(* IEC 61131-3 sources: 2026_Projet_YGO_ExcavatriceDragage/CODE_BACKUP/CODE_20260822_IntroductionTestCI/J_SUPERVISION/_TYPES/4_JOYSTICK_ACQUISITION, 9 files *)

(* ---- ST_AcquisitionInterPrg.st ---- *)
(* ═══════════════════════════════════════════════════════════════
   🧲 ST_AcquisitionInterPrg — Bus d'échange inter-PRG produit par PRG_02_Acquisition
   ───────────────────────────────────────────────────────────────
   🎯 Rôle : Encapsuler les mesures câbles/vitesses, les états joystick qualifiés,
      les positions M3 et les diagnostics DI publiés par PRG_02_Acquisition vers
      les consommateurs (PRG_03/04/05/07, FB_TroubleshootingView).
   📤 Producteur unique : PRG_02_Acquisition (VAR_OUTPUT Data : ST_AcquisitionInterPrg).
   📄 Doc : DOC/AF/AF_Partie-06_Acquisition_Qualification_IO_v2.3.md
   🔌 Architecture : Bus de données typé — encapsulation des échanges inter-PRG.
   ═══════════════════════════════════════════════════════════════ *)

TYPE ST_AcquisitionInterPrg :
STRUCT
    // === 🧲 Mesures câbles & vitesses treuils M1/M2 ===
    CablePosM1              : REAL; // 📏 Position cable M1 calibree (metres)
    CablePosM2              : REAL; // 📏 Position cable M2 calibree (metres)
    M1_Speed_Mps            : REAL; // 📏 Vitesse absolue M1 (m/s)
    M1_SignedSpeed_Mps      : REAL; // 📏 Vitesse signee M1 (+:Montee, -:Descente) (m/s)
    M1_SpeedValid           : BOOL; // 🟢 Validite mesure vitesse M1
    M2_Speed_Mps            : REAL; // 📏 Vitesse absolue M2 (m/s)
    M2_SignedSpeed_Mps      : REAL; // 📏 Vitesse signee M2 (+:Montee, -:Descente) (m/s)
    M2_SpeedValid           : BOOL; // 🟢 Validite mesure vitesse M2

    // === 🕹️ États joystick qualifiés ===
    JoystickDeadmanArmed    : BOOL; // 🔒 Homme-mort joystick arme (1=Arme)
    JoystickYNeutral        : BOOL; // 🟢 Axe Y joystick au neutre
    JoystickDirectionX      : INT;  // 🎯 Sens X demande (-1:Gauche, 0:Neutre, 1:Droite)
    JoystickSpeedPctX       : REAL; // 📈 Magnitude deviation axe X en % (0..100)
    JoystickXNeutral        : BOOL; // 🟢 Axe X joystick au neutre

    // === 🎯 Positions translation M3 (zones cumulatives + points exacts) ===
    TranslationPosTremie      : BOOL; // 📍 Zone Tremie (1=Present)
    TranslationPosPV          : BOOL; // 📍 Zone pre-ralentissement PV (1=Present)
    TranslationPosP2          : BOOL; // 📍 Zone P2 (1=Present)
    TranslationPosP1          : BOOL; // 📍 Zone P1 (1=Present)
    TranslationPosMaintenance : BOOL; // 📍 Zone Maintenance (1=Present)
    TranslationAtTremie       : BOOL; // 🎯 Position exacte Tremie (1=Atteint)
    TranslationAtPV           : BOOL; // 🎯 Position exacte PV (1=Atteint)
    TranslationAtP2           : BOOL; // 🎯 Position exacte P2 (1=Atteint)
    TranslationAtP1           : BOOL; // 🎯 Position exacte P1 (1=Atteint)
    TranslationAtMaintenance  : BOOL; // 🎯 Position exacte Maintenance (1=Atteint)
    M3_LimitSwitchFwd         : BOOL; // 🛡️ Fin de course avant M3 (1=Actionne)
    M3_LimitSwitchRev         : BOOL; // 🛡️ Fin de course arriere M3 (1=Actionne)
    M3_SensorWordIncoherent   : BOOL; // ❌ Incoherence detectee mot capteurs M3
    M3_SensorsWord             : BYTE; // 📊 Mot d'etat capteurs M3

    // === 🩺 Diagnostics modules DI & codeurs ===
    LocalDigitalIoOk         : BOOL; // 🟢 Module Local_Digital_IO OK
    Vh0800EndOk              : BOOL; // 🟢 Module VH_0800END OK
    Vh0808EtpOk              : BOOL; // 🟢 Module VH_0808ETP OK
    InputModuleFault         : BOOL; // ❌ Defaut sur au moins un module DI
    M1_EncoderIncoherent     : BOOL; // ❌ Mesure codeur M1 incoherente
    M2_EncoderIncoherent     : BOOL; // ❌ Mesure codeur M2 incoherente
    M1_EncoderFault          : BOOL; // ❌ Gate fiabilite M1 (NOT Available OR Incoherent, sans Homed)
    M2_EncoderFault          : BOOL; // ❌ Gate fiabilite M2 (NOT Available OR Incoherent, sans Homed)
    M1_HomedAndReliable      : BOOL; // ✅ Gate strict M3 M1 : dispo ET reference ET pas incoherent
    M2_HomedAndReliable      : BOOL; // ✅ Gate strict M3 M2 : dispo ET reference ET pas incoherent

    // === 🧪 Simulation & variateur M3 filtré ===
    WinchInputSourceChanged       : BOOL; // 🔀 Impulsion 1 cycle si source Winch bascule (IHM)
    M3_StatusWord_Filtered        : UINT; // 📊 Mot d'etat variateur M3 filtre (consommé PRG_05)
    M3_ActualFrequencyHz_Filtered : UINT; // 📊 Frequence reelle M3 filtree (consommé PRG_05)
END_STRUCT
END_TYPE

(* ---- ST_EncoderHMI.st ---- *)
(* ═══════════════════════════════════════════════════════════════
   🧲 ST_EncoderHMI — Données d'échange IHM pour les codeurs absolus
   ───────────────────────────────────────────────────────────────
   🎨 Destiné à l'affichage des informations et diagnostics des codeurs.
   ═══════════════════════════════════════════════════════════════ *)
TYPE ST_EncoderHMI :
STRUCT
    RawPos           : UDINT; (* 📊 Position brute lue sur le bus *)
    Alarms           : UINT;  (* ⚠️ Code d'alarme brut du codeur *)
    Warnings         : UINT;  (* 🟧 Code d'avertissement brut du codeur *)
    SlaveOperational : BOOL;  (* 📡 Esclave EtherCAT opérationnel *)
    PresetTriggerCmd : WORD;  (* 🎯 Commande de preset active *)
    PresetValueOut   : UDINT; (* 📐 Valeur de preset envoyée au codeur *)
    Error            : BOOL;  (* Codeur en défaut (liaison EtherCAT ou preset) *)
    ErrorId          : WORD;  (* ❌ Code défaut codeur *)

    (* 🎯 Homing — prise d'origine / référencement *)
    Homed                   : BOOL;             (* 🎯 Prise d'origine (Homing) validée *)
    HomingBusy              : BOOL;             (* ⏳ Référencement en cours *)
    HomingDone              : BOOL;             (* ✅ Pulse de référencement réussi *)
    HomingError             : BOOL;             (* Défaut de référencement *)
    HomingErrorId           : WORD;             (* ❌ Bitfield défaut homing *)
    HomingState             : E_State;          (* 🤖 État FB_Encoder_Homing *)
    HomingStateAtError      : E_State;          (* 🧭 État lors du défaut *)
    HomingSuspect           : BOOL;             (* ⚠️ Référence à confirmer *)
    HomingRefRaw            : UDINT;            (* 📐 Référence brute appliquée *)
END_STRUCT
END_TYPE

(* ---- ST_HardwareImage.st ---- *)
(* ═══════════════════════════════════════════════════════════════
   🏗️ ST_HardwareImage — Structure globale d'image matérielle (Frontière HwIn)
   ───────────────────────────────────────────────────────────────
   🎨 Agrège les 4 sous-domaines matériels : Winch, Translation, Operator, Machine.
   ═══════════════════════════════════════════════════════════════ *)
TYPE ST_HardwareImage :
STRUCT
    Winch       : ST_HwWinch;       (* Entrées brutes domaine Treuils M1/M2 + codeurs *)
    Translation : ST_HwTranslation; (* Entrées brutes domaine Translation M3 + variateur *)
    Operator    : ST_HwOperator;    (* Entrées brutes domaine Opérateur / Joystick / bus CAN *)
    Machine     : ST_HwMachine;     (* Entrées brutes domaine Sécurités/Communs Machine *)
END_STRUCT
END_TYPE

(* ---- ST_HwMachine.st ---- *)
(* ═══════════════════════════════════════════════════════════════
   🏗️ ST_HwMachine — Image matérielle brute des entrées communes Machine
   ───────────────────────────────────────────────────────────────
   🎨 Regroupe les signaux physiques d'entrée bruts communs à la machine.
   ═══════════════════════════════════════════════════════════════ *)
TYPE ST_HwMachine :
STRUCT
    PowerContactorEngaged_DI       : BOOL; (* Confirm. contacteur puissance engagé *)
    EmergencyChainClosed_DI        : BOOL; (* Boucle AU fermée (coup-de-poing + contact PLC) *)
    PhaseRotationOk_DI             : BOOL; (* Contrôle rotation phases élec. OK *)
    M1_M2_M3_BrakeThermalOk_DI     : BOOL; (* Thermique frein M1/M2/M3 commun OK *)
    M1_M2_KoboldBottomTouch_DI     : BOOL; (* Retour détecteur fond Kobold *)
    HydraulicThermalOk_DI          : BOOL; (* Thermique centrale hydraulique OK *)
    ConveyorInfeedReady_DI         : BOOL; (* Autorisation démarrage crible (dépôt gravats) *)
    HopperFull_OR_GateRaised_DI    : BOOL; (* : Trémie pleine OU grille levée — pas encore câblé électriquement,
                                               déclaré en avance (Device_IO_20260812). Aucun consommateur pour l'instant :
                                               l'interdiction translation M3→Trémie est une tâche à part, voir PLAN_TASK.md. *)
END_STRUCT
END_TYPE

(* ---- ST_HwOperator.st ---- *)
(* ═══════════════════════════════════════════════════════════════
   🏗️ ST_HwOperator — Image matérielle brute des entrées Opérateur / Joystick
   ───────────────────────────────────────────────────────────────
   🎨 Regroupe les signaux physiques d'entrée bruts du joystick CANopen JOY1.
   ═══════════════════════════════════════════════════════════════ *)
TYPE ST_HwOperator :
STRUCT
    JoyXRaw_ANA1      : INT;          (* Valeur brute analogique axe X (Translation) *)
    JoyYRaw_ANA2      : INT;          (* Valeur brute analogique axe Y (Levage) *)
    JoyBtnRaw         : BOOL;         (* Bouton brut joystick (Homme-Mort) *)
    CanBusState       : INT;          (* État bus CANopen (CANbus.GetBusState) *)
    JOY1_DeviceState  : DEVICE_STATE; (* État device JOY1 (GetDeviceState) *)
END_STRUCT
END_TYPE

(* ---- ST_JoystickChecklist.st ---- *)
(* ═══════════════════════════════════════════════════════════════
   🕹️ ST_JoystickChecklist — Diagnostic chronologique communication & prise en main Joystick
   ───────────────────────────────────────────────────────────────
   🎨 Permet de vérifier la chaîne Joystick (CANopen, Homme-mort, Neutre, Calibration).
   ═══════════════════════════════════════════════════════════════ *)
TYPE ST_JoystickChecklist :
STRUCT
    (* 1. Bus & Matériel *)
    Step1_CanBusActive           : BOOL; (* TRUE = Bus CANopen en état ACTIVE *)
    Step2_JoystickOperational    : BOOL; (* TRUE = Esclave JOY1 en état RUNNING *)

    (* 1bis. Entrées physiques directes HwIn *)
    HwIn_JoyBtnRaw_DI            : BOOL; (* Bouton brut homme-mort issu de HwIn.Operator *)
    NeutralXAct                  : BOOL; (* TRUE = Axe X au neutre (PRG_02_Acquisition.JoystickXNeutral) *)
    NeutralYAct                  : BOOL; (* TRUE = Axe Y au neutre (PRG_02_Acquisition.JoystickYNeutral) *)

    (* 2. Prise en main & Sécurité *)
    Step3_DeadmanPressed         : BOOL; (* TRUE = Bouton Homme-Mort appuyé *)
    Step4_NeutralAcquired        : BOOL; (* TRUE = Repassé par le neutre (autorisation mouvement) *)
    DeadmanArmed                 : BOOL; (* TRUE = Homme-Mort armé avec passage au neutre validé *)

    (* 3. Éligibilité globale *)
    AllConditionsMet             : BOOL; (* TRUE = Joystick prêt pour piloter un axe *)
    JoystickSelected             : BOOL; (* TRUE = Joystick maître sélectionné IHM *)
    SelJoystickWinch             : INT;  (* Sélection Treuil (0=Couplé M1+M2, 1=M1 seul, 2=M2 seul) *)

    (* 4. Mesures brutes & Filtrées *)
    RawX                         : INT;  (* Valeur brute axe X (0..10000) *)
    RawY                         : INT;  (* Valeur brute axe Y (0..10000) *)
    DeflectionX_Pct              : REAL; (* Déflexion signée X (%) *)
    DeflectionY_Pct              : REAL; (* Déflexion signée Y (%) *)
    DirectionX                   : INT;  (* Direction filtrée X (-1 / 0 / +1) *)
    DirectionY                   : INT;  (* Direction filtrée Y (-1 / 0 / +1) *)
END_STRUCT
END_TYPE

(* ---- ST_JoystickCmd.st ---- *)
(* ═══════════════════════════════════════════════════════════════
   🎮 ST_JoystickCmd — Commandes IHM pour le Joystick
   ═══════════════════════════════════════════════════════════════ *)
TYPE ST_JoystickCmd :
STRUCT
    BtnCalibrate : BOOL; (* 🎯 Demande de recalage au neutre *)
END_STRUCT
END_TYPE

(* ---- ST_JoystickHMI.st ---- *)
(* ═══════════════════════════════════════════════════════════════
   🕹️ ST_JoystickHMI — Données d'échange IHM pour le Joystick
   ───────────────────────────────────────────────────────────────
   📄 Structuration en Cmd / State , homogène avec ST_ModesHMI.
   Pas de Cfg (les vrais réglages de calibration vivent dans GVL_PERSISTENT, pas ici) ni de
   Bypass (concept absent de ce struct).
   ═══════════════════════════════════════════════════════════════ *)
TYPE ST_JoystickHMI :
STRUCT
    Cmd   : ST_JoystickCmd;
    State : ST_JoystickState;
END_STRUCT
END_TYPE

(* ---- ST_JoystickState.st ---- *)
(* ═══════════════════════════════════════════════════════════════
   🚦 ST_JoystickState — États et diagnostics IHM du Joystick
   ═══════════════════════════════════════════════════════════════ *)
TYPE ST_JoystickState :
STRUCT
    RawX         : INT;        (* 🕹️ Axe X brut du joystick (0..10000) *)
    RawY         : INT;        (* 🕹️ Axe Y brut du joystick (0..10000) *)
    RawButton    : BOOL;       (* 🔘 Bouton homme-mort brut *)
    AxisCmdX     : ST_Joystick_AxisCmd; (* ⚙️ Consigne d'axe X normalisée (sortie FB_Joystick) *)
    AxisCmdY     : ST_Joystick_AxisCmd; (* ⚙️ Consigne d'axe Y normalisée (sortie FB_Joystick) *)
    NeutralXAct  : INT;        (* 🎯 Neutre X calibré actuel (lecture seule) *)
    NeutralYAct  : INT;        (* 🎯 Neutre Y calibré actuel (lecture seule) *)
    DeadmanArmed : BOOL;       (* 🔫 Geste homme-mort armé (FB_Joystick.DeadmanArmed) *)
    AtNeutral    : BOOL;       (* : TRUE si les 2 axes sont en zone morte (position centrale) *)
    Online       : BOOL;       (* 📡 Liaison CAN joystick active *)
    Operational  : BOOL;       (* 🟢 Joystick opérationnel *)
    Error        : BOOL;       (* Joystick en défaut *)
    ErrorId      : WORD;       (* ❌ Code défaut joystick *)
END_STRUCT
END_TYPE
